// TIA Portal V15.1 export
// export: Created 2026-11-02T18:55:12.3319593Z, ExportSetting WithDefaults, DisplayName Totally Integrated Automation Portal, DisplayVersion V15.1, DisplayName TIA Portal Openness, DisplayVersion V15.1, DisplayName STEP 7 Professional, DisplayVersion V15.1, DisplayName WinCC Professional, DisplayVersion V15.1
VAR_GLOBAL   // PLC tag table "IO"
   PSH_101 AT %I0.0 : Bool;   // Scrubber high pressure
   LSH_102 AT %I0.1 : Bool;   // Scrubber high level
   LSHH_103 AT %I0.2 : Bool;   // Scrubber high-high level
   BR01_Run AT %I0.3 : Bool;   // BR01 run feedback
   S1_BR01_Start AT %I0.4 : Bool;   // BR01 START push button
   BR01_Fault AT %I0.5 : Bool;   // BR01 fault (lockout)
   S3_BR01_Stop AT %I0.6 : Bool;   // BR01 STOP push button
   S0_EStopStatus AT %I1.0 : Bool;   // E-STOP status (NC1)
   S2_FaultReset AT %I1.1 : Bool;   // FAULT RESET push button
   LSL_TK01 AT %I1.2 : Bool;   // TK01 low level
   LSL_TK02 AT %I1.3 : Bool;   // TK02 low level
   BR02_Run AT %I1.4 : Bool;   // BR02 run feedback
   BR02_Fault AT %I1.5 : Bool;   // BR02 fault (lockout)
   Rfuel2_BR02_DieselMode AT %I12.0 : Bool;   // BR02 diesel mode
   S4_BR01_Auto AT %I12.1 : Bool;   // BR01 AUTO/MAN selector (closed = AUTO)
   S5_BR02_Auto AT %I12.2 : Bool;   // BR02 AUTO/MAN selector (closed = AUTO)
   S6_BR02_Start AT %I12.3 : Bool;   // BR02 START push button
   S7_BR02_Stop AT %I12.4 : Bool;   // BR02 STOP push button
   BR01_TL_Cmd AT %Q0.0 : Bool;   // BR01 heat request (TL) + H1 1st stage lamp
   BR01_TR_Cmd AT %Q0.1 : Bool;   // BR01 2nd stage (TR) + H2 2nd stage lamp
   XV_401_Cmd AT %Q0.2 : Bool;   // XV-401 Flare SV (NO)
   XV_402_Cmd AT %Q0.3 : Bool;   // XV-402 Drain SV (NC)
   XV_403_Cmd AT %Q0.4 : Bool;   // XV-403 Suction SV (NC)
   BR02_L_Cmd AT %Q0.5 : Bool;   // BR02 start (L)
   BR02_T2_Cmd AT %Q0.6 : Bool;   // BR02 high fire (T2)
   BR02_Stage1Lamp_Cmd AT %Q0.7 : Bool;   // BR02 1st stage lamp H5
   BR02_Stage2Lamp_Cmd AT %Q1.0 : Bool;   // BR02 2nd stage lamp H6
   TE_501_Raw AT %IW96 : Int;   // TK01 inlet oil temperature
   TE_502_Raw AT %IW98 : Int;   // TK01 outlet oil temperature
   TE_503_Raw AT %IW100 : Int;   // TK02 inlet oil temperature
   TE_504_Raw AT %IW102 : Int;   // TK02 outlet oil temperature
END_VAR
